TYPE ST_TwinSAFE :
STRUCT
	TSafeIn			AT %I*	: TwinSafeOut_PlcIn;
	TSafeOut		AT %Q*	: TwinSafeIn_PlcOut;
	stSafetyIn		AT %I* 	: ST_SafeOut_PlcIn;
	stSafetyOut		AT %Q* 	: ST_SafeIn_PlcOut;	
END_STRUCT
END_TYPE

(* stored: Version 1.1.0.1, ProductVersion 3.1.4024.12
   DUT ST_TwinSAFE: Id {fbeb76a3-97f9-48e1-a517-9acb0dceeafb} *)
